(* IEC 61131-3 sources: volt/packages/volt-lsp-iec/test-corpus/lenze-mid/Device/Plc Logic/Application/A71_LocalSources, 2 files *)

(* ---- Scale_Offset_Dint.pou ---- *)
FUNCTION Scale_Offset_Dint
VAR_INPUT
	iX1 : DINT;
	iX2 : DINT;
	iY1 : DINT;
	iY2 : DINT;
	iXvalue : DINT;

END_VAR
VAR

END_VAR
VAR_OUTPUT
	oyValue_DI : DINT;
	oYValue_R : REAL;
	oPercentage_R : REAL;
	oPercentage_I : INT;
END_VAR

%LANGUAGE ST

END_FUNCTION

(* ---- POU_systemStart.pou ---- *)
PROGRAM POU_systemStart
VAR
END_VAR

%LANGUAGE LD
%NETWORK
ASSIGN(RAIL(), Q_SET => LST_General.FirstCycle);

END_PROGRAM
